// TIA Portal V20 export
// export: Created 2026-10-12T15:48:31.2157525Z, ExportSetting WithDefaults, DisplayName Totally Integrated Automation Portal, DisplayVersion V20, DisplayName TIA Portal Openness, DisplayVersion V20, DisplayName TIA Portal Teamcenter Gateway, DisplayVersion V20, DisplayName TIA Portal Version Control Interface, DisplayVersion V20, DisplayName SINAMICS Startdrive Advanced, DisplayVersion V20 SP1 Update 2, DisplayName SINAMICS Startdrive G110M, G120, G120C, G120D, G120P, G115D, DisplayVersion V20 SP1 Update 2, DisplayName SINAMICS Startdrive G130, G150, S120, S150, SINAMICS MV, G220, S200, S210, DisplayVersion V20 SP1 Update 2, DisplayName STEP 7 Professional, DisplayVersion V20, DisplayName STEP 7 Safety, DisplayVersion V20, DisplayName WinCC Basic/Comfort/Advanced, DisplayVersion V20, DisplayName WinCC Professional, DisplayVersion V20, DisplayName WinCC Unified, DisplayVersion V20
FUNCTION "FRK_ConfigRevision" : UDInt   // FC23, SCL
{ S7_Optimized_Access := 'TRUE' }
VERSION : 0.1
// Core 3.10.2: deterministic typed walk, one bounded response window.
//  Static facets carry no write capability. Every reused slot is cleared.
// stored: AutoNumber true, IsIECCheckEnabled false, SetENOAutomatically false, UDAEnableTagReadback false
   VAR_INPUT
      Previous : UDInt;
   END_VAR
   VAR_TEMP
      Stamp : DTL;
      ResultCode : Int;
      Generation : ULInt;
   END_VAR
BEGIN

   #FRK_ConfigRevision := #Previous + 1;
   #ResultCode := RD_SYS_T(OUT => #Stamp);
   IF #ResultCode = 0 THEN
       #Generation := LDT_TO_ULINT(DTL_TO_LDT(#Stamp)) / ULINT#1000000;
       #FRK_ConfigRevision := ULINT_TO_UDINT(#Generation MOD ULINT#4294967296);
   END_IF;
   IF #FRK_ConfigRevision = #Previous THEN
       #FRK_ConfigRevision := #Previous + 1;
   END_IF;
   IF #FRK_ConfigRevision = 0 THEN
       #FRK_ConfigRevision := 1;
   END_IF;
END_FUNCTION
